(* Single Solid Attenuator (SATT) filter stack (L2SI compact, 4 stacks
   of 8 filters): single-axis mover via FB_PositionStateND (states OUT,
   FILTER1..FILTER8). Not a PMPS state mover; only RTD reactive-temp
   fault thresholds and a "device moving" fast fault. Per-cycle transmission
   from filter material/thickness and beam energy. Deps injected via FB_Init. *)
{attribute 'call_after_init'}
FUNCTION_BLOCK FB_SXR_SATT_Stage
VAR_INPUT
    (* Per-filter material / thickness table. Used by the transmission
       calculation. Index 1 corresponds to FILTER1 (which is the
       state at slot 2 in astPositionState, since OUT lives at slot 1
       in E_SXR_SATT_Position). *)
    {attribute 'pytmc' := 'pv: FILTERS'}
    arrFilters : ARRAY[1..8] OF ST_SATT_Filter;
END_VAR
VAR_OUTPUT
    fTemp1                    : LREAL;
    fTemp2                    : LREAL;
    bIsStationary             : BOOL;
    bError                    : BOOL;
    // The current position state as an enum.
    {attribute 'pytmc' := '
        pv: STATE:GET
        io: i
    '}
    eEnumGet : E_SXR_SATT_Position;
    {attribute 'pytmc' := '
        pv: MATERIAL
        io: i
    '}
    sActiveFilterMaterial     : STRING;

    {attribute 'pytmc' := '
        pv: THICKNESS
        io: i
        field: EGU um
    '}
    fActiveFilterThickness_um : LREAL;

    {attribute 'pytmc' := '
        pv: TRANSMISSION
        io: i
        field: DESC Filter transmission
    '}
    fTransmission             : LREAL;
    fActiveFilterDensity      : LREAL;
    fActiveFilterAtomicMass   : LREAL;
    fAbsorptionConstant       : LREAL;

    iFilterIndex              : INT := 0;
END_VAR
VAR
    (* State-enum bridge bound to FB_PositionStateND's REFERENCE TO UINT
       param via the shared UINT base. EPICS owns it through the pytmc
       pragma; PLC code must go through the EnumSet property instead of
       touching it directly. *)
    // Set this to a non-unknown value to request a new move.
    {attribute 'pytmc' := '
        pv: STATE:SET
        io: io
    '}
    eEnumSet : E_SXR_SATT_Position;

    fbStates : FB_PositionStateND(
        aiMotionStage        := aiMotionStage,
        astPositionState     := astPositionState,
        nActiveMotorCount    := 1,
        eEnumSet             := eEnumSet,
        eEnumGet             := eEnumGet,
        bEnableMotion        := bEnableMotion,
        eMotionRequestPolicy := E_MotionRequestPolicy.INTERRUPT
    );

    fbAtomicMass               : FB_AtomicMass;
    fbAttenuatorElementDensity : FB_AttenuatorElementDensity;

    (* EL3202-0020: 0.01 deg C per digit. Vetoed when the stage is in
       OUT (no filter in beam, no temperature to monitor). *)
    {attribute 'pytmc' := 'pv: RTD:1'}
    fbRTD_1 : FB_CC_TempSensor := (fResolution := 0.01);
    {attribute 'pytmc' := 'pv: RTD:2'}
    fbRTD_2 : FB_CC_TempSensor := (fResolution := 0.01);

    bFileReaderBusy       : REFERENCE TO BOOL;
    (* Per-cycle JSON DB read for the currently active filter's
       PMPS state, just to pull the reactive temp setpoint into
       astPickedDB[1].stReactiveParams.nTempSP. Not a PMPS BPTM
       participant; just borrows the DB pipeline. *)
    fbReadPMPSDB : FB_JsonDocToSafeBP;
    astPickedDB  : ARRAY[1..1] OF ST_DbStateParams;

    (* "Device is moving" fast fault. Raised while the Y motor is
       moving or while we are sitting in UNKNOWN. *)
    fbFF : FB_FastFault := (
        i_Desc       := 'Device is moving',
        i_TypeCode   := E_MotionFFType.DEVICE_MOVE,
        i_xAutoReset := TRUE
    );

    (* REFERENCE TO backing fields populated by FB_Init. *)
    {attribute 'no_copy'}
    aiMotionStage    : REFERENCE TO ARRAY[1..MotionConstants.MAX_STATE_MOTORS] OF I_MotionStage;
    {attribute 'no_copy'}
    astPositionState : REFERENCE TO ARRAY[1..MotionConstants.MAX_STATE_MOTORS]
                                          OF ARRAY[1..GeneralConstants.MAX_STATES] OF ST_PositionState;
    {attribute 'no_copy'}
    fbFFHWO          : REFERENCE TO FB_HardwareFFOutput;
    sDeviceName      : STRING;
    (* PMPS DB key for the RTD reactive-temperature read. The filters are not real PMPS states,
        so this device-level key names the DB entry to pull the reactive temp setpoint from.
    *)
    RTDPMPSState     : STRING;
    bEnableMotion    : BOOL := TRUE;
END_VAR

(* Nil-ref guards: every REFERENCE TO backing field must be bound. *)
IF NOT __ISVALIDREF(aiMotionStage)
   OR NOT __ISVALIDREF(astPositionState)
   OR NOT __ISVALIDREF(fbFFHWO) THEN
    RETURN;
END_IF

fbStates();

(* Filter index is offset by one because E_SXR_SATT_Position.OUT
   occupies slot 1 and FILTER1..FILTER8 occupy slots 2..9. *)
iFilterIndex := UINT_TO_INT(eEnumGet) - 1;

IF iFilterIndex >= 1 AND iFilterIndex <= 8 THEN
    sActiveFilterMaterial     := arrFilters[iFilterIndex].sFilterMaterial;
    fActiveFilterThickness_um := arrFilters[iFilterIndex].fFilterThickness_um;

    fbAtomicMass(
        sName  := sActiveFilterMaterial,
        fValue => fActiveFilterAtomicMass
    );
    fbAttenuatorElementDensity(
        sName    := sActiveFilterMaterial,
        fDensity => fActiveFilterDensity
    );

    fAbsorptionConstant := F_CalculateAbsorptionConstant(
        sElement      := sActiveFilterMaterial,
        fEnergyEV     := PMPS_GVL.stCurrentBeamParameters.neV,
        fDensity_gm3  := fActiveFilterDensity,
        fAtomicWeight := fActiveFilterAtomicMass,
        bError        => bError
    );
    fTransmission := F_CalculateTransmission(
        fAbsorptionConstant := fAbsorptionConstant,
        fThickness_in_m     := fActiveFilterThickness_um * 1.0E-6
    );
ELSE
    sActiveFilterMaterial     := '';
    fActiveFilterThickness_um := 0.0;
    fAbsorptionConstant       := 0.0;
    fActiveFilterDensity      := 0.0;
    fActiveFilterAtomicMass   := 0.0;
    fTransmission             := 1.0;
END_IF

(* "Device is moving" fault: stationary AND known position. Reads the
   motor's NC status through the I_MotionStage interface; aiMotionStage
   was nil-guarded above so slot 1 deref is safe. *)
bIsStationary := NOT aiMotionStage[1].Axis.Status.Moving;
fbFF(
    i_DevName  := sDeviceName,
    i_xOK      := bIsStationary AND eEnumGet <> E_SXR_SATT_Position.UNKNOWN,
    io_fbFFHWO := fbFFHWO
);

(* The RTD reactive-temperature read is keyed on the device-level
   RTDPMPSState (the filters are not real PMPS states, so no per-
   filter key is scanned). The named DB entry must exist; the
   temperature field may be blank. *)
astPickedDB[1].sPmpsState := RTDPMPSState;

fbReadPMPSDB(
    bExecute    := NOT bFileReaderBusy,
    jsonDoc     := PMPS_GVL.BP_jsonDoc,
    sDeviceName := sDeviceName,
    arrStates   := astPickedDB,
    io_fbFFHWO  := fbFFHWO
);

fbRTD_1(
    fFaultThreshold := astPickedDB[1].stReactiveParams.nTempSP,
    sDevName        := sDeviceName,
    bVeto           := eEnumGet = E_SXR_SATT_Position.OUT,
    io_fbFFHWO      := fbFFHWO
);
fTemp1 := fbRTD_1.fTemp;

fbRTD_2(
    fFaultThreshold := astPickedDB[1].stReactiveParams.nTempSP,
    sDevName        := sDeviceName,
    bVeto           := eEnumGet = E_SXR_SATT_Position.OUT,
    io_fbFFHWO      := fbFFHWO
);
fTemp2 := fbRTD_2.fTemp;

(* Auto-fired after FB_Init. fbStates' inline-init ran first and
   forwarded nil refs, so this re-supplies the now-valid refs via
   fbStates.CallAfterInitStateMover, running the Core / ND wiring chain. *)
{attribute 'call_after_init'}
METHOD CallAfterInit
THIS^.fbStates.CallAfterInitStateMover(
    aiMotionStage         := aiMotionStage,
    astPositionState      := astPositionState,
    nActiveMotorCount     := 1,
    eEnumSet              := eEnumSet,
    eEnumGet              := eEnumGet,
    bEnableMotion         := bEnableMotion,
    eMotionRequestPolicy  := E_MotionRequestPolicy.INTERRUPT,
);
END_METHOD

(* Stores all FB_Init inputs into instance fields. Every input is
   REFERENCE TO and is REF= bound for the lifetime of the FB.
   Inline-init of fbStates above runs first, capturing the FB_Init
   params at construction time; this method then records the same
   references on THIS^ for body-side use and live caller writes. *)
{attribute 'analysis' := '-33'}
METHOD FB_Init : BOOL
VAR_INPUT
    bInitRetains     : BOOL;
    bInCopyCode      : BOOL;
    aiMotionStage    : REFERENCE TO ARRAY[1..MotionConstants.MAX_STATE_MOTORS] OF I_MotionStage;
    astPositionState : REFERENCE TO ARRAY[1..MotionConstants.MAX_STATE_MOTORS]
                                          OF ARRAY[1..GeneralConstants.MAX_STATES] OF ST_PositionState;
    bFileReaderBusy       : REFERENCE TO BOOL;
    fbFFHWO          : REFERENCE TO FB_HardwareFFOutput;
    sDeviceName      : STRING;
    RTDPMPSState     : STRING;
END_VAR
THIS^.aiMotionStage    REF= aiMotionStage;
THIS^.astPositionState REF= astPositionState;
THIS^.fbFFHWO          REF= fbFFHWO;
THIS^.bFileReaderBusy 	REF=bFileReaderBusy;
THIS^.sDeviceName      := sDeviceName;
THIS^.RTDPMPSState     := RTDPMPSState;
END_METHOD

(* Current position state. Read-only; written by the state mover. *)
PROPERTY EnumGet : E_SXR_SATT_Position
GET
EnumGet := eEnumGet;
END_GET
END_PROPERTY

(* Request a new move, e.g. `fbSATT.EnumSet := E_SXR_SATT_Position.FILTER1;`.
   The state mover consumes and clears the request. *)
PROPERTY EnumSet : E_SXR_SATT_Position
GET
EnumSet := eEnumSet;
END_GET
SET
eEnumSet := EnumSet;
END_SET
END_PROPERTY

END_FUNCTION_BLOCK

(* stored: Version 1.1.0.1
   POU FB_SXR_SATT_Stage: Id {7fb611c7-2215-4e8f-8a28-e51a98acae9a}, SpecialFunc None
   Method CallAfterInit: Id {7fb611c8-2215-4e8f-8a28-e51a98acae9b}
   Method FB_init: Id {7fb611c9-2215-4e8f-8a28-e51a98acae9c}
   Property EnumGet: Id {176f7c09-c56c-42e7-b20a-6b0da2f13387}
   Get Get: Id {63dfefc0-6337-4760-bade-4056669f937c}
   Property EnumSet: Id {b7616b49-7981-48ca-aef7-a43b09424e67}
   Get Get: Id {5da9a31e-56f3-40ba-b74f-384ca8163935}
   Set Set: Id {60c02dbe-7fb8-4781-abdf-ebabce3efb88} *)
